(* IEC 61131-3 sources: nautilus/examples/spatial-rig, 3 files *)

(* ---- types.st ---- *)
(* One UDT per kind of physical prop on the rig. A 3D or AR scene binds a
   whole asset by its tag name (T101, P101, XV101) and reads the members,
   so these structs are the contract between the rig and the scene file.
   A root .st with no PROGRAM is a library: `type: Tank` in the manifest
   resolves against it. *)

TYPE
  Tank : STRUCT
    Level : REAL;   (* % *)
    TempC : REAL;
    HH    : BOOL;   (* limit bits the alarm rules claim *)
    LL    : BOOL;
  END_STRUCT;

  Motor : STRUCT
    Run   : BOOL;   (* command *)
    Running : BOOL; (* feedback *)
    Fault : BOOL;
    Speed : REAL;   (* % *)
    Hours : REAL;
  END_STRUCT;

  Valve : STRUCT
    Cmd    : REAL;  (* % open command *)
    Pos    : REAL;  (* % open feedback *)
    Fault  : BOOL;  (* position disagrees with command *)
  END_STRUCT;

  (* A UDT of UDTs: a transfer skid is a pump and a valve. The 3D scene's
     assembly kind binds one Skid tag and its parts read the members
     (SK101.Pump, SK101.Valve) — docs/design/spatial-hmi.md §3d. Fault is
     the skid's own bit, because alarm rules match one level of members. *)
  Skid : STRUCT
    Pump  : Motor;
    Valve : Valve;
    Fault : BOOL;
  END_STRUCT;
END_TYPE

(* ---- control.st ---- *)
PROGRAM Control
(* The rig's control logic: P-101 fills T-101 between two levels, XV-101
   follows the operator's demand, and the limit bits the alarms claim. *)
VAR_EXTERNAL
    T101 : Tank;
    P101 : Motor;
    XV101 : Valve;
    SK101 : Skid;
    SK102 : Skid;
    Demand : REAL;
    StartLevel : REAL;
    StopLevel : REAL;
    LevelHH : REAL;
    LevelLL : REAL;
    ControlDtS : REAL;
END_VAR

(* pump seal-in: start below StartLevel, stop above StopLevel, never on a fault *)
IF P101.Fault THEN
    P101.Run := FALSE;
ELSIF T101.Level < StartLevel THEN
    P101.Run := TRUE;
ELSIF T101.Level > StopLevel THEN
    P101.Run := FALSE;
END_IF;

IF P101.Running THEN
    P101.Hours := P101.Hours + ControlDtS / 3600.0;
END_IF;

XV101.Cmd := LIMIT(0.0, Demand, 100.0);
XV101.Fault := ABS(XV101.Cmd - XV101.Pos) > 10.0;

T101.HH := T101.Level > LevelHH;
T101.LL := T101.Level < LevelLL;

(* transfer skids: the duty skid runs while the drain passes flow, its valve
   opens with its pump; the standby takes over when the duty pump faults *)
SK101.Pump.Run := XV101.Pos > 5.0 AND NOT SK101.Pump.Fault;
SK102.Pump.Run := XV101.Pos > 5.0 AND SK101.Pump.Fault AND NOT SK102.Pump.Fault;
IF SK101.Pump.Run THEN
    SK101.Valve.Cmd := 100.0;
ELSE
    SK101.Valve.Cmd := 0.0;
END_IF;
IF SK102.Pump.Run THEN
    SK102.Valve.Cmd := 100.0;
ELSE
    SK102.Valve.Cmd := 0.0;
END_IF;
SK101.Fault := SK101.Pump.Fault;
SK102.Fault := SK102.Pump.Fault;
END_PROGRAM

(* ---- sim.st ---- *)
PROGRAM Sim
(* Stands in for the field. The props on the office rig are dumb objects;
   this task gives them a moving process, plus fault-injection switches so
   an AR panel has alarms and bad states to show on demand. *)
VAR_EXTERNAL
    T101 : Tank;
    P101 : Motor;
    XV101 : Valve;
    SK101 : Skid;
    SK102 : Skid;
    SimDtS : REAL;
    InjectPumpFault : BOOL;
    InjectValveStick : BOOL;
END_VAR
VAR CONSTANT
    CapacityL  : REAL := 100.0;   (* small, so a fill/drain cycle is ~2 min *)
    PumpMaxLps : REAL := 1.0;
    DrainMaxLps : REAL := 0.8;
    ValveRatePctS : REAL := 20.0;  (* stroke speed *)
    PumpRampPctS : REAL := 25.0;
END_VAR
VAR
    inLps : REAL;
    outLps : REAL;
    step : REAL;
END_VAR

P101.Fault := InjectPumpFault;
P101.Running := P101.Run AND NOT P101.Fault;
IF P101.Running THEN
    P101.Speed := MIN(P101.Speed + PumpRampPctS * SimDtS, 100.0);
ELSE
    P101.Speed := MAX(P101.Speed - PumpRampPctS * SimDtS, 0.0);
END_IF;

(* the valve strokes toward its command unless it is stuck *)
IF NOT InjectValveStick THEN
    step := ValveRatePctS * SimDtS;
    XV101.Pos := XV101.Pos + LIMIT(-step, XV101.Cmd - XV101.Pos, step);
END_IF;

inLps := P101.Speed / 100.0 * PumpMaxLps;
outLps := XV101.Pos / 100.0 * DrainMaxLps * SQRT(T101.Level / 100.0);
T101.Level := LIMIT(0.0, T101.Level + (inLps - outLps) * SimDtS / CapacityL * 100.0, 100.0);
T101.TempC := 20.0 + 0.05 * P101.Speed;

(* the transfer skids: the injected pump fault trips the duty skid too, so
   the standby has something to take over from *)
SK101.Pump.Fault := InjectPumpFault;
SK101.Pump.Running := SK101.Pump.Run AND NOT SK101.Pump.Fault;
IF SK101.Pump.Running THEN
    SK101.Pump.Speed := MIN(SK101.Pump.Speed + PumpRampPctS * SimDtS, 100.0);
ELSE
    SK101.Pump.Speed := MAX(SK101.Pump.Speed - PumpRampPctS * SimDtS, 0.0);
END_IF;
step := ValveRatePctS * SimDtS;
SK101.Valve.Pos := SK101.Valve.Pos + LIMIT(-step, SK101.Valve.Cmd - SK101.Valve.Pos, step);

SK102.Pump.Running := SK102.Pump.Run AND NOT SK102.Pump.Fault;
IF SK102.Pump.Running THEN
    SK102.Pump.Speed := MIN(SK102.Pump.Speed + PumpRampPctS * SimDtS, 100.0);
ELSE
    SK102.Pump.Speed := MAX(SK102.Pump.Speed - PumpRampPctS * SimDtS, 0.0);
END_IF;
SK102.Valve.Pos := SK102.Valve.Pos + LIMIT(-step, SK102.Valve.Cmd - SK102.Valve.Pos, step);
END_PROGRAM
